(* IEC 61131-3 sources: beedance/embedded/bench/st, 2 files *)

(* ---- calc.st ---- *)
(* The arithmetic workload of the embedded benchmark: a loop of integer and
   real operations, the instruction dispatch and arithmetic of each engine
   with no function block or I/O. acc ends at 303 every scan. *)
PROGRAM Main
VAR
    i : DINT;
    acc : DINT;
    x : REAL;
END_VAR
acc := 0;
FOR i := 1 TO 100 DO
    acc := acc + (i * 3) MOD 7;
    x := x * 0.5 + 1.0;
END_FOR;
END_PROGRAM

(* ---- plc.st ---- *)
(* The PLC program of the esp32hw firmware: a TON that restarts itself,
   so %QX0.0 pulses once every 1 s and two scans. On the device's clock the
   pulses come 1020 ms apart at 10 ms scans; embedded/esp32hw checks them
   against the host's clock. *)
PROGRAM Main
VAR
    t : TON;
    pulses : DINT;
    pulse AT %QX0.0 : BOOL;
END_VAR
t(IN := NOT t.Q, PT := T#1s);
IF t.Q THEN
    pulses := pulses + 1;
END_IF;
pulse := t.Q;
END_PROGRAM
